Universal Robots PolyScope program: new.urp

Program new (installation=default directory=/programs createdIn=5.23.0 lastSavedIn=5.23.0 robotSerialNumber=20245590068)
Calibrated DH parameters: a=[0.00013, -0.03651, -0.389144, 0.000102, 0.000008, 0]; d=[0.162613, 192.230671, -179.915756, -12.181517, 0.099698, 0.099535]; alpha=[1.57038, 0.002205, 0.004138, 1.570804, -1.571025, 0]; deltaTheta=[-0.000001, 1.484886, 4.928506, -0.130209, 0, 0]
InitVariablesNode
Robot Program (runOnlyOnce=false)
  Placeholder
